SYSTEM System (* System Configuration *)
  (* Standard: 61499-1 *)
  (* Version 0.0, 7/14/2023, Cheyan, Schneider Electric *)
  {SET_ATTRIBUTE(System.Device.FolderPath, EcoRT_0)}
  APPLICATION APP1
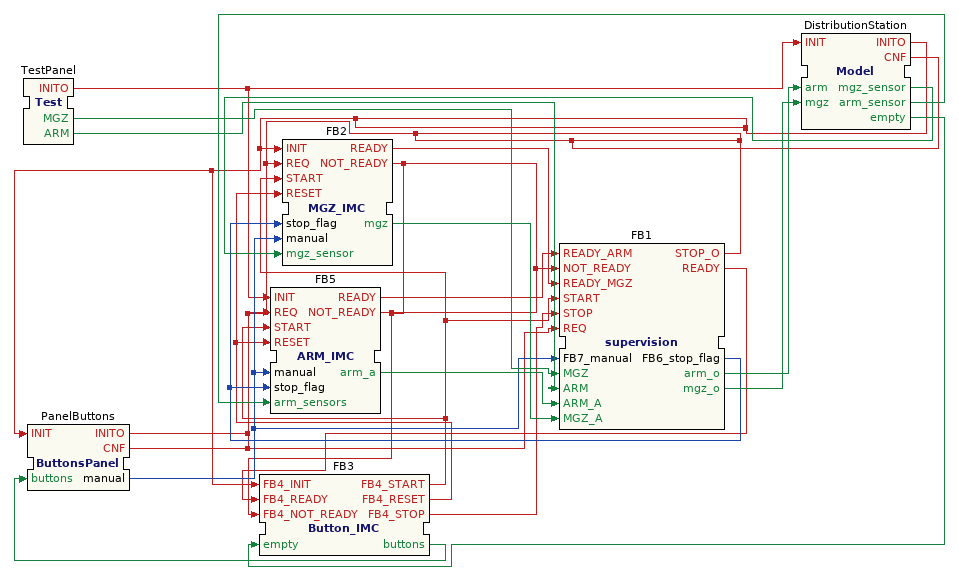
    (* HMI *)
    (* Supervision *)
    (* CONTROL *)
    (* MODEL *)
    FBS
      TestPanel : Test;
      DistributionStation : Model;
      PanelButtons : ButtonsPanel;
      FB2 : MGZ_IMC;
      FB1 : supervision;
      FB5 : ARM_IMC;
      FB3 : Button_IMC;
    END_FBS
    EVENT_CONNECTIONS
      TestPanel.INITO TO DistributionStation.INIT;
      DistributionStation.INITO TO PanelButtons.INIT;
      DistributionStation.INITO TO FB2.INIT;
      PanelButtons.INITO TO FB2.REQ;
      FB1.STOP_O TO FB2.REQ;
      FB5.READY TO FB1.READY_ARM;
      FB5.NOT_READY TO FB1.NOT_READY;
      FB2.READY TO FB1.READY_MGZ;
      FB2.NOT_READY TO FB1.NOT_READY;
      TestPanel.INITO TO FB5.INIT;
      DistributionStation.CNF TO FB5.REQ;
      PanelButtons.INITO TO FB5.REQ;
      FB1.STOP_O TO FB5.REQ;
      DistributionStation.INITO TO FB3.FB4_INIT;
      FB1.READY TO FB3.FB4_READY;
      FB5.NOT_READY TO FB3.FB4_NOT_READY;
      FB2.NOT_READY TO FB3.FB4_NOT_READY;
      FB3.FB4_START TO FB2.START;
      FB3.FB4_START TO FB1.START;
      FB3.FB4_START TO FB5.START;
      FB3.FB4_RESET TO FB2.RESET;
      FB3.FB4_RESET TO FB5.RESET;
      FB3.FB4_STOP TO FB1.STOP;
      PanelButtons.CNF TO FB5.REQ;
      PanelButtons.CNF TO FB2.REQ;
      PanelButtons.CNF TO FB1.REQ;
    END_CONNECTIONS
    DATA_CONNECTIONS
      PanelButtons.manual TO FB1.FB7_manual;
      FB1.FB6_stop_flag TO FB2.stop_flag;
      PanelButtons.manual TO FB5.manual;
      FB1.FB6_stop_flag TO FB5.stop_flag;
      PanelButtons.manual TO FB2.manual;
    END_CONNECTIONS
    ADAPTER_CONNECTIONS
      TestPanel.MGZ TO FB1.MGZ;
      TestPanel.ARM TO FB1.ARM;
      FB5.arm_a TO FB1.ARM_A;
      FB2.mgz TO FB1.MGZ_A;
      DistributionStation.mgz_sensor TO FB2.mgz_sensor;
      FB1.arm_o TO DistributionStation.arm;
      FB1.mgz_o TO DistributionStation.mgz;
      DistributionStation.arm_sensor TO FB5.arm_sensors;
      DistributionStation.empty TO FB3.empty;
      FB3.buttons TO PanelButtons.buttons;
    END_CONNECTIONS
  END_APPLICATION
  DEVICE EcoRT_0 : Soft_dPAC
    RESOURCE RES0 : EMB_RES_ECO
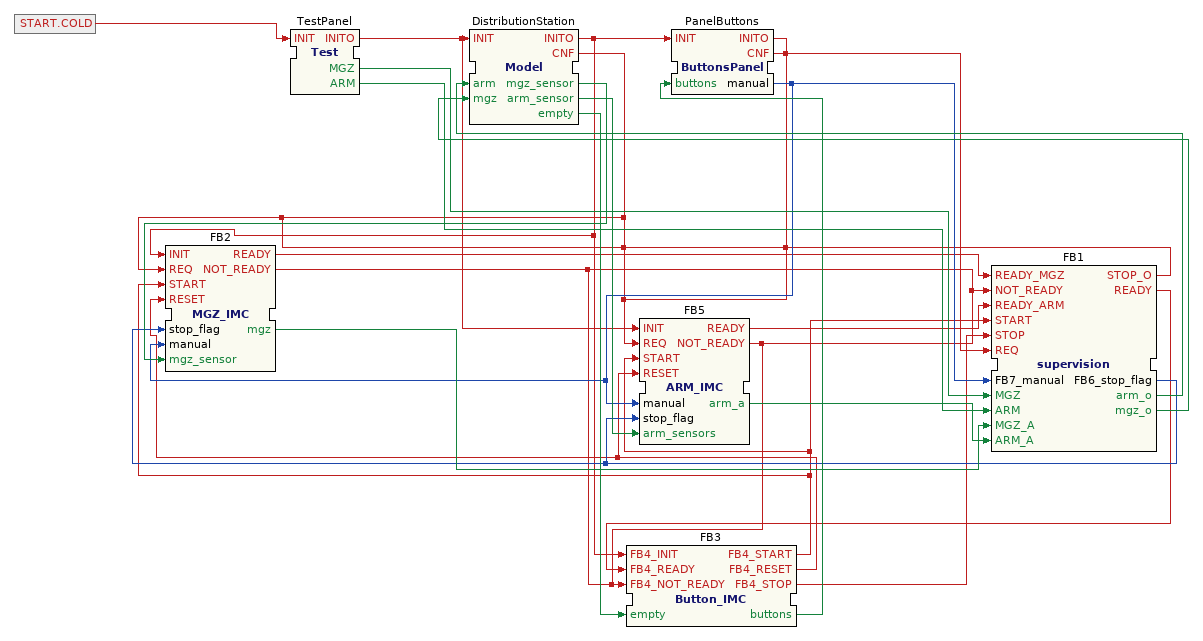
      FBS
        TestPanel : Test;
        DistributionStation : Model;
        PanelButtons : ButtonsPanel;
        FB2 : MGZ_IMC;
        FB1 : supervision;
        FB5 : ARM_IMC;
        FB3 : Button_IMC;
      END_FBS
      EVENT_CONNECTIONS
        TestPanel.INITO TO DistributionStation.INIT;
        START.COLD TO TestPanel.INIT;
        DistributionStation.INITO TO PanelButtons.INIT;
        DistributionStation.INITO TO FB2.INIT;
        PanelButtons.INITO TO FB2.REQ;
        FB1.STOP_O TO FB2.REQ;
        FB2.READY TO FB1.READY_MGZ;
        FB2.NOT_READY TO FB1.NOT_READY;
        FB5.READY TO FB1.READY_ARM;
        FB5.NOT_READY TO FB1.NOT_READY;
        TestPanel.INITO TO FB5.INIT;
        DistributionStation.CNF TO FB5.REQ;
        PanelButtons.INITO TO FB5.REQ;
        FB1.STOP_O TO FB5.REQ;
        DistributionStation.INITO TO FB3.FB4_INIT;
        FB1.READY TO FB3.FB4_READY;
        FB5.NOT_READY TO FB3.FB4_NOT_READY;
        FB2.NOT_READY TO FB3.FB4_NOT_READY;
        FB3.FB4_START TO FB2.START;
        FB3.FB4_START TO FB1.START;
        FB3.FB4_START TO FB5.START;
        FB3.FB4_RESET TO FB2.RESET;
        FB3.FB4_RESET TO FB5.RESET;
        FB3.FB4_STOP TO FB1.STOP;
        PanelButtons.CNF TO FB5.REQ;
        PanelButtons.CNF TO FB2.REQ;
        PanelButtons.CNF TO FB1.REQ;
      END_CONNECTIONS
      DATA_CONNECTIONS
        PanelButtons.manual TO FB1.FB7_manual;
        FB1.FB6_stop_flag TO FB2.stop_flag;
        PanelButtons.manual TO FB5.manual;
        FB1.FB6_stop_flag TO FB5.stop_flag;
        PanelButtons.manual TO FB2.manual;
      END_CONNECTIONS
      ADAPTER_CONNECTIONS
        TestPanel.MGZ TO FB1.MGZ;
        TestPanel.ARM TO FB1.ARM;
        FB2.mgz TO FB1.MGZ_A;
        DistributionStation.mgz_sensor TO FB2.mgz_sensor;
        FB1.arm_o TO DistributionStation.arm;
        FB1.mgz_o TO DistributionStation.mgz;
        FB5.arm_a TO FB1.ARM_A;
        DistributionStation.arm_sensor TO FB5.arm_sensors;
        DistributionStation.empty TO FB3.empty;
        FB3.buttons TO PanelButtons.buttons;
      END_CONNECTIONS
    END_RESOURCE
  END_DEVICE
  MAPPINGS
    APP1.TestPanel ON EcoRT_0.RES0;
    APP1.DistributionStation ON EcoRT_0.RES0;
    APP1.PanelButtons ON EcoRT_0.RES0;
    APP1.FB2 ON EcoRT_0.RES0;
    APP1.FB1 ON EcoRT_0.RES0;
    APP1.FB5 ON EcoRT_0.RES0;
    APP1.FB3 ON EcoRT_0.RES0;
  END_MAPPINGS
END_SYSTEM
